FUNCTION_BLOCK DistributingSequence (* Basic Function Block Type *)
  (* Standard: 61499-2 *)
  (* Version 0.0, 11/16/2026, Sandeep Patil, Flexbridge AB, Template *)
  PACKAGE Flexbridge.FestoMPS400;
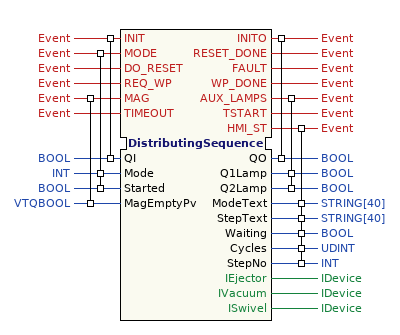
  EVENT_INPUT
    INIT WITH QI; (* Initialisation request *)
    MODE WITH Mode, Started; (* Station mode changed (StationMode) *)
    DO_RESET; (* Run the reset sequence (StationMode) *)
    REQ_WP; (* Request one workpiece (Testing, or the HMI button) *)
    MAG WITH MagEmptyPv; (* Magazine sensor changed *)
    TIMEOUT; (* Ejection pulse time over (EjectTimer) *)
  END_EVENT
  EVENT_OUTPUT
    INITO WITH QO; (* Initialisation confirm *)
    RESET_DONE; (* Reset sequence finished (StationMode) *)
    FAULT; (* Stopped on a device fault (StationMode) *)
    WP_DONE; (* Workpiece handed over (Testing) *)
    AUX_LAMPS WITH Q1Lamp, Q2Lamp; (* Console lamps Q1 and Q2 *)
    TSTART; (* Start the ejection pulse timer *)
    HMI_ST WITH ModeText, StepText, Waiting, Cycles, StepNo; (* State for the HMI *)
  END_EVENT
  VAR_INPUT
    QI : BOOL; (* Input event qualifier *)
    Mode : INT; (* Station mode: 0 = wait for RESET, 1 = resetting, 2 = wait for START, 3 = started *)
    Started : BOOL; (* Station started: requests are accepted *)
    MagEmptyPv : VTQBOOL; (* B4 magazine empty *)
  END_VAR
  VAR_OUTPUT
    QO : BOOL; (* Output event qualifier *)
    Q1Lamp : BOOL; (* Lamp Q1: waiting, magazine empty *)
    Q2Lamp : BOOL; (* Lamp Q2: not used *)
    ModeText : STRING[40]; (* Station mode as text *)
    StepText : STRING[40]; (* Current step as text (number and name) *)
    Waiting : BOOL; (* Waiting for workpieces (magazine empty) *)
    Cycles : UDINT; (* Workpieces handed over since start-up *)
    StepNo : INT; (* Current step number *)
  END_VAR
  PLUGS
    IEjector : IDevice;
    IVacuum : IDevice;
    ISwivel : IDevice;
  END_PLUGS
  VAR
    Done : BOOL; (* The current step has reached its target *)
    Fault : BOOL; (* A device needs Rearm, or is not program local when it must be *)
    InCycle : BOOL; (* Parking belongs to a workpiece cycle (else to the reset sequence) *)
    Accept : BOOL; (* A workpiece request is accepted (station started) *)
    RdySwivel : BOOL; (* Swivel has sent CNF_READY: its owner has initialised *)
    AdpSwivel : BOOL; (* Swivel taken over at start-up, or the reset sequence has run *)
    TrySwivel : INT; (* Program-local requests sent to Swivel at start-up *)
  END_VAR
  EC_STATES
    START; (* Initial state *)
    INIT_S : algInit, algModeText, -> AUX_LAMPS, -> HMI_ST, -> INITO;
    S_IDLE : algModeText, algIdle -> HMI_ST;
    IDLE_W; (* Idle: wait for RESET (reset sequence) or a workpiece request *)
    M_IDLE : algModeText -> HMI_ST;
    S_R_SEL : algModeText, algS_R_SEL -> HMI_ST, -> IEjector.REQ_PROGLOCALSEL, -> IVacuum.REQ_PROGLOCALSEL, -> ISwivel.REQ_PROGLOCALSEL, -> AUX_LAMPS;
    C_R_SEL : algC_R_SEL;
    W_R_SEL; (* Wait: Reset: owners to program *)
    S_R_HOME : algModeText, algS_R_HOME -> HMI_ST, -> IVacuum.REQ_CMD, -> IEjector.REQ_CMD;
    C_R_HOME : algC_R_HOME;
    W_R_HOME; (* Wait: Reset: ejector home *)
    S_P_MAG : algModeText, algS_P_MAG -> HMI_ST, -> ISwivel.REQ_CMD;
    C_P_MAG : algC_P_MAG;
    W_P_MAG; (* Wait: Park: swivel to magazine *)
    S_P_OFF : algModeText, algS_P_OFF -> HMI_ST, -> ISwivel.REQ_CMD;
    C_P_OFF : algC_P_OFF;
    W_P_OFF; (* Wait: Park: off the magazine *)
    S_P_STOP : algModeText, algS_P_STOP -> HMI_ST, -> ISwivel.REQ_CMD;
    S_R_DONE : algModeText, algS_R_DONE -> HMI_ST, -> RESET_DONE;
    Q_CHK : algQ_CHK;
    Q_NOSTART : algModeText -> HMI_ST;
    S_C_MAG : algModeText, algS_C_MAG -> HMI_ST, -> AUX_LAMPS;
    W_C_MAG; (* Wait: magazine empty *)
    S_C_PUSH : algModeText, algS_C_PUSH -> HMI_ST, -> IEjector.REQ_CMD;
    C_C_PUSH : algC_C_PUSH;
    W_C_PUSH; (* Wait: Push workpiece out *)
    S_C_BACK : algModeText, algS_C_BACK -> HMI_ST, -> IEjector.REQ_CMD;
    C_C_BACK : algC_C_BACK;
    W_C_BACK; (* Wait: Ejector back home *)
    S_C_TOMAG : algModeText, algS_C_TOMAG -> HMI_ST, -> ISwivel.REQ_CMD;
    C_C_TOMAG : algC_C_TOMAG;
    W_C_TOMAG; (* Wait: Swivel to magazine *)
    S_C_GRIP : algModeText, algS_C_GRIP -> HMI_ST, -> IVacuum.REQ_CMD;
    C_C_GRIP : algC_C_GRIP;
    W_C_GRIP; (* Wait: Vacuum on, wait gripped *)
    S_C_TODOWN : algModeText, algS_C_TODOWN -> HMI_ST, -> ISwivel.REQ_CMD;
    C_C_TODOWN : algC_C_TODOWN;
    W_C_TODOWN; (* Wait: Swivel to Testing *)
    S_C_REL : algModeText, algS_C_REL -> HMI_ST, -> IVacuum.REQ_CMD, -> TSTART;
    W_C_REL; (* Wait: ejection pulse *)
    K_C_REL : algK_C_REL;
    S_C_VACOFF : algModeText, algS_C_VACOFF -> HMI_ST, -> IVacuum.REQ_CMD;
    S_C_DONE : algModeText, algS_C_DONE -> HMI_ST, -> AUX_LAMPS, -> WP_DONE;
    FAULT_S : algModeText, algFault -> HMI_ST, -> AUX_LAMPS, -> FAULT; (* Fault: RESET restarts the reset sequence after Rearm on the faceplate *)
    SR_Swivel : algRdySwivel; (* Swivel ready before INIT *)
    TR_Swivel : algRdySwivel;
    TK_Swivel; (* Start-up takeover of Swivel *)
    TS_Swivel : algTkSelSwivel -> ISwivel.REQ_PROGLOCALSEL;
    TC_Swivel : algTkCmdSwivel -> ISwivel.REQ_CMD;
  END_STATES
  EC_TRANSITIONS
    START TO INIT_S := INIT;
    INIT_S TO S_IDLE := 1;
    S_IDLE TO TK_Swivel := 1;
    IDLE_W TO INIT_S := INIT;
    IDLE_W TO M_IDLE := MODE;
    M_IDLE TO IDLE_W := 1;
    IDLE_W TO S_R_SEL := DO_RESET;
    IDLE_W TO Q_CHK := REQ_WP;
    S_R_SEL TO C_R_SEL := 1;
    C_R_SEL TO FAULT_S := Fault;
    C_R_SEL TO S_R_HOME := NOT Fault AND Done;
    C_R_SEL TO W_R_SEL := NOT Fault AND NOT Done;
    W_R_SEL TO C_R_SEL := IEjector.CNF_STATUS OR IEjector.CNF_READY OR IVacuum.CNF_STATUS OR IVacuum.CNF_READY OR ISwivel.CNF_STATUS OR ISwivel.CNF_READY;
    S_R_HOME TO C_R_HOME := 1;
    C_R_HOME TO FAULT_S := Fault;
    C_R_HOME TO S_P_MAG := NOT Fault AND Done;
    C_R_HOME TO W_R_HOME := NOT Fault AND NOT Done;
    W_R_HOME TO C_R_HOME := IEjector.CNF_STATUS OR IEjector.CNF_READY OR IVacuum.CNF_STATUS OR IVacuum.CNF_READY OR ISwivel.CNF_STATUS OR ISwivel.CNF_READY;
    S_P_MAG TO C_P_MAG := 1;
    C_P_MAG TO FAULT_S := Fault;
    C_P_MAG TO S_P_OFF := NOT Fault AND Done;
    C_P_MAG TO W_P_MAG := NOT Fault AND NOT Done;
    W_P_MAG TO C_P_MAG := IEjector.CNF_STATUS OR IEjector.CNF_READY OR IVacuum.CNF_STATUS OR IVacuum.CNF_READY OR ISwivel.CNF_STATUS OR ISwivel.CNF_READY;
    S_P_OFF TO C_P_OFF := 1;
    C_P_OFF TO FAULT_S := Fault;
    C_P_OFF TO S_P_STOP := NOT Fault AND Done;
    C_P_OFF TO W_P_OFF := NOT Fault AND NOT Done;
    W_P_OFF TO C_P_OFF := IEjector.CNF_STATUS OR IEjector.CNF_READY OR IVacuum.CNF_STATUS OR IVacuum.CNF_READY OR ISwivel.CNF_STATUS OR ISwivel.CNF_READY;
    S_P_STOP TO S_C_DONE := InCycle;
    S_P_STOP TO S_R_DONE := NOT InCycle;
    S_R_DONE TO IDLE_W := 1;
    Q_CHK TO Q_NOSTART := NOT Accept;
    Q_NOSTART TO IDLE_W := 1;
    Q_CHK TO FAULT_S := Accept AND Fault;
    Q_CHK TO S_C_MAG := Accept AND NOT Fault;
    S_C_MAG TO S_C_PUSH := NOT Waiting;
    S_C_MAG TO W_C_MAG := Waiting;
    W_C_MAG TO S_C_MAG := MAG;
    S_C_PUSH TO C_C_PUSH := 1;
    C_C_PUSH TO FAULT_S := Fault;
    C_C_PUSH TO S_C_BACK := NOT Fault AND Done;
    C_C_PUSH TO W_C_PUSH := NOT Fault AND NOT Done;
    W_C_PUSH TO C_C_PUSH := IEjector.CNF_STATUS OR IEjector.CNF_READY OR IVacuum.CNF_STATUS OR IVacuum.CNF_READY OR ISwivel.CNF_STATUS OR ISwivel.CNF_READY;
    S_C_BACK TO C_C_BACK := 1;
    C_C_BACK TO FAULT_S := Fault;
    C_C_BACK TO S_C_TOMAG := NOT Fault AND Done;
    C_C_BACK TO W_C_BACK := NOT Fault AND NOT Done;
    W_C_BACK TO C_C_BACK := IEjector.CNF_STATUS OR IEjector.CNF_READY OR IVacuum.CNF_STATUS OR IVacuum.CNF_READY OR ISwivel.CNF_STATUS OR ISwivel.CNF_READY;
    S_C_TOMAG TO C_C_TOMAG := 1;
    C_C_TOMAG TO FAULT_S := Fault;
    C_C_TOMAG TO S_C_GRIP := NOT Fault AND Done;
    C_C_TOMAG TO W_C_TOMAG := NOT Fault AND NOT Done;
    W_C_TOMAG TO C_C_TOMAG := IEjector.CNF_STATUS OR IEjector.CNF_READY OR IVacuum.CNF_STATUS OR IVacuum.CNF_READY OR ISwivel.CNF_STATUS OR ISwivel.CNF_READY;
    S_C_GRIP TO C_C_GRIP := 1;
    C_C_GRIP TO FAULT_S := Fault;
    C_C_GRIP TO S_C_TODOWN := NOT Fault AND Done;
    C_C_GRIP TO W_C_GRIP := NOT Fault AND NOT Done;
    W_C_GRIP TO C_C_GRIP := IEjector.CNF_STATUS OR IEjector.CNF_READY OR IVacuum.CNF_STATUS OR IVacuum.CNF_READY OR ISwivel.CNF_STATUS OR ISwivel.CNF_READY;
    S_C_TODOWN TO C_C_TODOWN := 1;
    C_C_TODOWN TO FAULT_S := Fault;
    C_C_TODOWN TO S_C_REL := NOT Fault AND Done;
    C_C_TODOWN TO W_C_TODOWN := NOT Fault AND NOT Done;
    W_C_TODOWN TO C_C_TODOWN := IEjector.CNF_STATUS OR IEjector.CNF_READY OR IVacuum.CNF_STATUS OR IVacuum.CNF_READY OR ISwivel.CNF_STATUS OR ISwivel.CNF_READY;
    S_C_REL TO W_C_REL := 1;
    W_C_REL TO S_C_VACOFF := TIMEOUT;
    W_C_REL TO K_C_REL := IEjector.CNF_STATUS OR IEjector.CNF_READY OR IVacuum.CNF_STATUS OR IVacuum.CNF_READY OR ISwivel.CNF_STATUS OR ISwivel.CNF_READY;
    K_C_REL TO FAULT_S := Fault;
    K_C_REL TO W_C_REL := NOT Fault;
    S_C_VACOFF TO S_P_MAG := 1;
    S_C_DONE TO IDLE_W := 1;
    FAULT_S TO IDLE_W := 1;
    START TO SR_Swivel := ISwivel.CNF_READY;
    SR_Swivel TO START := 1;
    IDLE_W TO TR_Swivel := ISwivel.CNF_READY;
    TR_Swivel TO TK_Swivel := 1;
    IDLE_W TO TK_Swivel := ISwivel.CNF_STATUS;
    TK_Swivel TO TS_Swivel := NOT AdpSwivel AND RdySwivel AND NOT ISwivel.ProgLocal AND TrySwivel < 3;
    TK_Swivel TO TC_Swivel := NOT AdpSwivel AND RdySwivel AND ISwivel.ProgLocal AND (ISwivel.Status.value = 1 OR ISwivel.Status.value = 2);
    TK_Swivel TO IDLE_W := NOT (NOT AdpSwivel AND RdySwivel AND NOT ISwivel.ProgLocal AND TrySwivel < 3) AND NOT (NOT AdpSwivel AND RdySwivel AND ISwivel.ProgLocal AND (ISwivel.Status.value = 1 OR ISwivel.Status.value = 2));
    TS_Swivel TO IDLE_W := 1;
    TC_Swivel TO IDLE_W := 1;
  END_TRANSITIONS
  ALGORITHM algModeText IN ST: (* Station mode as text *)
CASE Mode OF
    0: ModeText := 'Wait for RESET';
    1: ModeText := 'Resetting';
    2: ModeText := 'Wait for START';
    3: ModeText := 'Started';
ELSE
    ModeText := 'Unknown mode';
END_CASE;
  END_ALGORITHM
  ALGORITHM algInit IN ST: (* Idle; lamps Q1 and Q2 off *)
QO := QI;
StepNo := 0; StepText := '0 Idle';
Waiting := FALSE; Q1Lamp := FALSE; Q2Lamp := FALSE;
InCycle := FALSE; Done := FALSE; Fault := FALSE;
Cycles := 0;
AdpSwivel := FALSE; TrySwivel := 0;
  END_ALGORITHM
  ALGORITHM algIdle IN ST: (* Idle *)
StepNo := 0; StepText := '0 Idle';
  END_ALGORITHM
  ALGORITHM algS_R_SEL IN ST: (* Reset: owners to program *)
StepNo := 10; StepText := '10 Reset: owners to program';
IEjector.ProgLocalSel := TRUE;
IVacuum.ProgLocalSel := TRUE;
ISwivel.ProgLocalSel := TRUE;
InCycle := FALSE; Waiting := FALSE; Q1Lamp := FALSE;
AdpSwivel := TRUE;
  END_ALGORITHM
  ALGORITHM algC_R_SEL IN ST: (* Check: Reset: owners to program *)
Fault := IEjector.NeedReset OR IVacuum.NeedReset OR ISwivel.NeedReset;
Done := IEjector.ProgLocal AND IVacuum.ProgLocal AND ISwivel.ProgLocal;
  END_ALGORITHM
  ALGORITHM algS_R_HOME IN ST: (* Reset: ejector home *)
StepNo := 11; StepText := '11 Reset: ejector home';
IVacuum.Lsp.value := 0;
IEjector.Lsp.value := 2;
  END_ALGORITHM
  ALGORITHM algC_R_HOME IN ST: (* Check: Reset: ejector home *)
Fault := IEjector.NeedReset OR IVacuum.NeedReset OR ISwivel.NeedReset;
Done := IEjector.Status.value = 2;
  END_ALGORITHM
  ALGORITHM algS_P_MAG IN ST: (* Park: swivel to magazine *)
StepNo := 20; StepText := '20 Park: swivel to magazine';
ISwivel.Lsp.value := 2;
  END_ALGORITHM
  ALGORITHM algC_P_MAG IN ST: (* Check: Park: swivel to magazine *)
Fault := IEjector.NeedReset OR IVacuum.NeedReset OR ISwivel.NeedReset;
Done := ISwivel.Status.value = 2;
  END_ALGORITHM
  ALGORITHM algS_P_OFF IN ST: (* Park: off the magazine *)
StepNo := 21; StepText := '21 Park: off the magazine';
ISwivel.Lsp.value := 1;
  END_ALGORITHM
  ALGORITHM algC_P_OFF IN ST: (* Check: Park: off the magazine *)
Fault := IEjector.NeedReset OR IVacuum.NeedReset OR ISwivel.NeedReset;
Done := ISwivel.Status.value <> 2;
  END_ALGORITHM
  ALGORITHM algS_P_STOP IN ST: (* Park: swivel stopped *)
StepNo := 22; StepText := '22 Park: swivel stopped';
ISwivel.Lsp.value := 0;
  END_ALGORITHM
  ALGORITHM algS_R_DONE IN ST: (* Reset done *)
StepNo := 12; StepText := '12 Reset done';
  END_ALGORITHM
  ALGORITHM algQ_CHK IN ST: (* Workpiece request: accept only when started and all devices ready *)
Accept := Started;
Fault := IEjector.NeedReset OR IVacuum.NeedReset OR ISwivel.NeedReset OR NOT (IEjector.ProgLocal AND IVacuum.ProgLocal AND ISwivel.ProgLocal);
IF NOT Accept THEN
    StepText := '0 Idle: press START first';
END_IF;
  END_ALGORITHM
  ALGORITHM algS_C_MAG IN ST: (* Cycle: wait while the magazine is empty *)
InCycle := TRUE;
Waiting := MagEmptyPv.value;
Q1Lamp := Waiting;
IF Waiting THEN
    StepNo := 31; StepText := '31 Wait: magazine empty';
ELSE
    StepNo := 31; StepText := '31 Magazine: workpiece there';
END_IF;
  END_ALGORITHM
  ALGORITHM algS_C_PUSH IN ST: (* Push workpiece out *)
StepNo := 32; StepText := '32 Push workpiece out';
IEjector.Lsp.value := 1;
  END_ALGORITHM
  ALGORITHM algC_C_PUSH IN ST: (* Check: Push workpiece out *)
Fault := IEjector.NeedReset OR IVacuum.NeedReset OR ISwivel.NeedReset;
Done := IEjector.Status.value = 1;
  END_ALGORITHM
  ALGORITHM algS_C_BACK IN ST: (* Ejector back home *)
StepNo := 33; StepText := '33 Ejector back home';
IEjector.Lsp.value := 2;
  END_ALGORITHM
  ALGORITHM algC_C_BACK IN ST: (* Check: Ejector back home *)
Fault := IEjector.NeedReset OR IVacuum.NeedReset OR ISwivel.NeedReset;
Done := IEjector.Status.value = 2;
  END_ALGORITHM
  ALGORITHM algS_C_TOMAG IN ST: (* Swivel to magazine *)
StepNo := 34; StepText := '34 Swivel to magazine';
ISwivel.Lsp.value := 2;
  END_ALGORITHM
  ALGORITHM algC_C_TOMAG IN ST: (* Check: Swivel to magazine *)
Fault := IEjector.NeedReset OR IVacuum.NeedReset OR ISwivel.NeedReset;
Done := ISwivel.Status.value = 2;
  END_ALGORITHM
  ALGORITHM algS_C_GRIP IN ST: (* Vacuum on, wait gripped *)
StepNo := 35; StepText := '35 Vacuum on, wait gripped';
IVacuum.Lsp.value := 1;
  END_ALGORITHM
  ALGORITHM algC_C_GRIP IN ST: (* Check: Vacuum on, wait gripped *)
Fault := IEjector.NeedReset OR IVacuum.NeedReset OR ISwivel.NeedReset;
Done := IVacuum.Status.value = 1;
  END_ALGORITHM
  ALGORITHM algS_C_TODOWN IN ST: (* Swivel to Testing *)
StepNo := 36; StepText := '36 Swivel to Testing';
ISwivel.Lsp.value := 1;
  END_ALGORITHM
  ALGORITHM algC_C_TODOWN IN ST: (* Check: Swivel to Testing *)
Fault := IEjector.NeedReset OR IVacuum.NeedReset OR ISwivel.NeedReset;
Done := ISwivel.Status.value = 1;
  END_ALGORITHM
  ALGORITHM algS_C_REL IN ST: (* Ejection pulse *)
StepNo := 37; StepText := '37 Release: ejection pulse';
IVacuum.Lsp.value := 2;
  END_ALGORITHM
  ALGORITHM algK_C_REL IN ST: (* Fault check while the pulse runs *)
Fault := IEjector.NeedReset OR IVacuum.NeedReset OR ISwivel.NeedReset;
  END_ALGORITHM
  ALGORITHM algS_C_VACOFF IN ST: (* Vacuum off *)
StepNo := 38; StepText := '38 Vacuum off';
IVacuum.Lsp.value := 0;
  END_ALGORITHM
  ALGORITHM algS_C_DONE IN ST: (* Cycle done: handed over *)
StepNo := 40; StepText := '40 Cycle done: handed over';
Cycles := Cycles + 1;
InCycle := FALSE; Waiting := FALSE; Q1Lamp := FALSE;
  END_ALGORITHM
  ALGORITHM algFault IN ST: (* Device fault: stop here, report to StationMode *)
StepNo := 99;
IF IEjector.NeedReset THEN
    StepText := '99 FAULT: Rearm Ejector';
ELSIF IVacuum.NeedReset THEN
    StepText := '99 FAULT: Rearm Vacuum';
ELSIF ISwivel.NeedReset THEN
    StepText := '99 FAULT: Rearm Swivel';
ELSE
    StepText := '99 FAULT: owner not program';
END_IF;
InCycle := FALSE; Waiting := FALSE; Q1Lamp := FALSE;
  END_ALGORITHM
  ALGORITHM algRdySwivel IN ST: (* Swivel has reported ready *)
RdySwivel := TRUE;
  END_ALGORITHM
  ALGORITHM algTkSelSwivel IN ST: (* Start-up: ask Swivel for program local *)
ISwivel.ProgLocalSel := TRUE;
TrySwivel := TrySwivel + 1;
  END_ALGORITHM
  ALGORITHM algTkCmdSwivel IN ST: (* Start-up: command the end position Swivel reports (it does not move) *)
ISwivel.Lsp.value := ISwivel.Status.value;
AdpSwivel := TRUE;
  END_ALGORITHM
END_FUNCTION_BLOCK
